TYPE ST_EL18x9 :
STRUCT
	
	State	AT %I*: UINT;
	i_ch1	AT %I*: BOOL;
	i_ch2	AT %I*: BOOL;
	i_ch3	AT %I*: BOOL;
	i_ch4	AT %I*: BOOL;
	i_ch5	AT %I*: BOOL;
	i_ch6	AT %I*: BOOL;
	i_ch7	AT %I*: BOOL;
	i_ch8	AT %I*: BOOL;
	
	i_ch9	AT %I*: BOOL;
	i_ch10	AT %I*: BOOL;
	i_ch11	AT %I*: BOOL;
	i_ch12	AT %I*: BOOL;
	i_ch13	AT %I*: BOOL;
	i_ch14	AT %I*: BOOL;
	i_ch15	AT %I*: BOOL;
	i_ch16	AT %I*: BOOL;
	
END_STRUCT
END_TYPE

(* stored: Version 1.1.0.1, ProductVersion 3.1.4024.12
   DUT ST_EL18x9: Id {dc4638ec-c66e-4410-8f4e-f0d9f097e07b} *)
